Fanuc KAREL source: kc00044.KL

-- PROVISIONAL review KL for V940-1; original PC SHA256 2f0432e54f59d2172199a955005e92e58bcefa207e87a3d0b1a28d8b0fce0474
-- Incomplete behavior may be omitted. Consult companion uncertainty JSON. Do not deploy.
PROGRAM KC00044
%NOLOCKGROUP
BEGIN
  -- V9_ZERO_TABLE_METADATA_HINT layout=0002_ascii; no indexed target words; source/name/runtime held
  -- UNRESOLVED_PC offsets 5-39; opcodes 27,22,22,22,22,22,31
  -- UNRESOLVED_PC offsets 44-48; opcodes 7F
END KC00044
